(* IEC 61131-3 sources: plcassist-cli/packages/volt-lsp-iec/test-corpus/lenze-mid/Device/Plc Logic/Application/Library Manager/CAA Async Manager, 30 files *)

(* ---- RSHANDLING.gvl ---- *)
VAR_GLOBAL
	G_JOBCLASS : JobClass;
END_VAR

(* ---- VERSIONCONSTANTS.gvl ---- *)
VAR_GLOBAL
	GC_BYVERSION : BYTE := 1;
	GC_BYVERSION_1 : BYTE := 0;
END_VAR

(* ---- _JOBABORT.fun ---- *)
FUNCTION _JOBABORT : ERROR
VAR_INPUT
	HJOB : CAA.HANDLE;
END_VAR
END_FUNCTION

(* ---- _JOBCLOSE.fun ---- *)
FUNCTION _JOBCLOSE : ERROR
VAR_INPUT
	HJOB : CAA.HANDLE;
END_VAR
END_FUNCTION

(* ---- _JOBEXECUTE.fun ---- *)
FUNCTION _JOBEXECUTE : ERROR
VAR_INPUT
	HJOB : CAA.HANDLE;
END_VAR
END_FUNCTION

(* ---- _JOBGETID.fun ---- *)
FUNCTION _JOBGETID : UDINT
VAR_INPUT
	HJOB : CAA.HANDLE;
	PEERROR : POINTER TO ERROR;
END_VAR
END_FUNCTION

(* ---- _JOBGETNUMOFJOBS.fun ---- *)
FUNCTION _JOBGETNUMOFJOBS : ERROR
VAR_IN_OUT
	NUMOFJOBS : ASM_CURRENT_MAX;
	NUMOFWORKERS : ASM_CURRENT_MAX;
END_VAR
END_FUNCTION

(* ---- _JOBGETPARAMS.fun ---- *)
FUNCTION _JOBGETPARAMS : CAA.PVOID
VAR_INPUT
	HJOB : CAA.HANDLE;
	PEERROR : POINTER TO ERROR;
END_VAR
END_FUNCTION

(* ---- _JOBGETSTATE.fun ---- *)
FUNCTION _JOBGETSTATE : ERROR
VAR_INPUT
	HJOB : CAA.HANDLE;
	PSTATEJOB : POINTER TO ASM_STATE;
END_VAR
END_FUNCTION

(* ---- _JOBOPEN.fun ---- *)
FUNCTION _JOBOPEN : CAA.HANDLE
VAR_INPUT
	UDIID : UDINT;
	PEERROR : POINTER TO ERROR;
END_VAR
END_FUNCTION

(* ---- _JOBOPENEX.fun ---- *)
FUNCTION _JOBOPENEX : CAA.HANDLE
VAR_INPUT
	UDIID : UDINT;
	PPARAMS : CAA.PVOID;
	PEERROR : POINTER TO ERROR;
END_VAR
END_FUNCTION

(* ---- _JOBRESET.fun ---- *)
FUNCTION _JOBRESET : ERROR
VAR_INPUT
	HJOB : CAA.HANDLE;
END_VAR
END_FUNCTION

(* ---- _JOBSETSTATE.fun ---- *)
FUNCTION _JOBSETSTATE : ERROR
VAR_INPUT
	HJOB : CAA.HANDLE;
	STATEJOB : ASM_STATE;
END_VAR
END_FUNCTION

(* ---- _WORKERREGISTER.fun ---- *)
FUNCTION _WORKERREGISTER : ERROR
VAR_INPUT
	UDIID : UDINT;
	PWITF : POINTER TO ASM_IWORKER;
END_VAR
END_FUNCTION

(* ---- _WORKERUNREGISTER.fun ---- *)
FUNCTION _WORKERUNREGISTER : ERROR
VAR_INPUT
	UDIID : UDINT;
END_VAR
END_FUNCTION

(* ---- GETSUPPLIERVERSION.fun ---- *)
FUNCTION GETSUPPLIERVERSION : WORD
END_FUNCTION

(* ---- JOBABORT.fun ---- *)
FUNCTION JOBABORT : ERROR
VAR_INPUT
	HJOB : CAA.HANDLE;
END_VAR
END_FUNCTION

(* ---- JOBCLOSE.fun ---- *)
FUNCTION JOBCLOSE : ERROR
VAR_INPUT
	HJOB : CAA.HANDLE;
END_VAR
END_FUNCTION

(* ---- JOBEXECUTE.fun ---- *)
FUNCTION JOBEXECUTE : ERROR
VAR_INPUT
	HJOB : CAA.HANDLE;
END_VAR
END_FUNCTION

(* ---- JOBGETID.fun ---- *)
FUNCTION JOBGETID : UDINT
VAR_INPUT
	HJOB : CAA.HANDLE;
	PEERROR : POINTER TO ERROR;
END_VAR
END_FUNCTION

(* ---- JOBGETNUMOFJOBS.fun ---- *)
FUNCTION JOBGETNUMOFJOBS : ERROR
VAR_INPUT
	NUMOFJOBS : POINTER TO ASM_CURRENT_MAX;
	NUMOFWORKERS : POINTER TO ASM_CURRENT_MAX;
END_VAR
END_FUNCTION

(* ---- JOBGETPARAMS.fun ---- *)
FUNCTION JOBGETPARAMS : CAA.PVOID
VAR_INPUT
	HJOB : CAA.HANDLE;
	PEERROR : POINTER TO ERROR;
END_VAR
END_FUNCTION

(* ---- JOBGETSTATE.fun ---- *)
FUNCTION JOBGETSTATE : ERROR
VAR_INPUT
	HJOB : CAA.HANDLE;
	PSTATEJOB : POINTER TO STATE;
END_VAR
END_FUNCTION

(* ---- JOBOPEN.fun ---- *)
FUNCTION JOBOPEN : CAA.HANDLE
VAR_INPUT
	UDIID : UDINT;
	PEERROR : POINTER TO ERROR;
END_VAR
END_FUNCTION

(* ---- JOBOPENEX.fun ---- *)
FUNCTION JOBOPENEX : CAA.HANDLE
VAR_INPUT
	UDIID : UDINT;
	PPARAMS : CAA.PVOID;
	PEERROR : POINTER TO ERROR;
END_VAR
END_FUNCTION

(* ---- JOBRESET.fun ---- *)
FUNCTION JOBRESET : ERROR
VAR_INPUT
	HJOB : CAA.HANDLE;
END_VAR
END_FUNCTION

(* ---- JOBSETSTATE.fun ---- *)
FUNCTION JOBSETSTATE : ERROR
VAR_INPUT
	HJOB : CAA.HANDLE;
	STATEJOB : ASM_STATE;
END_VAR
END_FUNCTION

(* ---- WORKERREGISTER.fun ---- *)
FUNCTION WORKERREGISTER : ERROR
VAR_INPUT
	UDIID : UDINT;
	PWITF : POINTER TO ASM_IWORKER;
END_VAR
END_FUNCTION

(* ---- WORKERUNREGISTER.fun ---- *)
FUNCTION WORKERUNREGISTER : ERROR
VAR_INPUT
	UDIID : UDINT;
END_VAR
END_FUNCTION

(* ---- JOBCLASS.fb ---- *)
FUNCTION_BLOCK JOBCLASS EXTENDS RSMClass
END_FUNCTION_BLOCK

METHOD CLOSE : RSM.ERROR
VAR_INPUT
	HHANDLE : CAA.HANDLE;
END_VAR
END_METHOD
